Universal Robots URScript: T013_zai-org_GLM-4.7-FP8_edit_perf_rep1.urscript

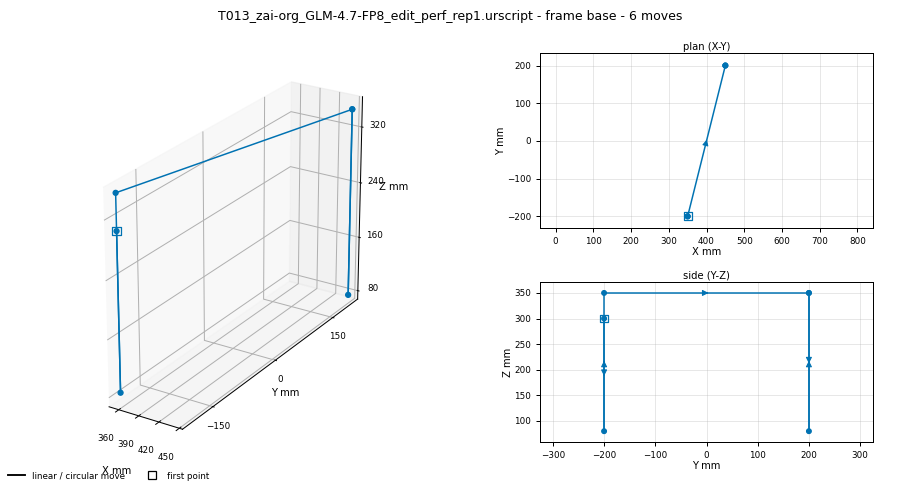
[picture p0: tool path of T013_zai-org_GLM-4.7-FP8_edit_perf_rep1.urscript in frame base, 6 of 8 moves have a stored position in this frame; points joined in program order, loops and branches not executed]
# Task: T013 — Collaborative suction palletizing — light boxes (Optimized)
# Generated by ENFIELD IR→URScript Translator
# Operating mode: collaborative | Max TCP speed: 0.250 m/s
# Robot: ur5e
#
# WARNING: This is auto-generated code for SIMULATION ONLY.
# Do NOT deploy to a physical robot without safety review.

def task_T013():
  # [0] E-Stop verify
  # E-Stop safety check (hardware-enforced on UR controller)
  if (get_digital_in(0) == True):
    popup("E-Stop active — aborting program.", error=True)
    halt
  end

  # [1] Home (Optimized: Increased joint velocity/acceleration)
  movej([0.0000, -1.5708, 1.5708, -1.5708, -1.5708, 0.0000], a=2.0000, v=1.5000)

  # [2] Above staging (Optimized: Max TCP speed, increased blend radius)
  movel(p[0.350000, -0.200000, 0.300000, 0.0000, 3.1416, 0.0000], a=1.2000, v=0.2500, r=0.0500)

  # [3] Descend to pick (Optimized: Slightly faster approach, no blend for precision)
  movel(p[0.350000, -0.200000, 0.080000, 0.0000, 3.1416, 0.0000], a=0.8000, v=0.1500, r=0.0000)

  # [4] Suction ON
  # set_tool (suction): {'vacuum_kpa': -40.0, 'state': 1.0}
  set_digital_out(0, True)

  # [5] Vacuum settle (Optimized: Reduced settle time for light payload)
  sleep(0.1000)

  # [6] Lift (Optimized: Max TCP speed, increased blend radius)
  movel(p[0.350000, -0.200000, 0.350000, 0.0000, 3.1416, 0.0000], a=1.2000, v=0.2500, r=0.0500)

  # [7] Transit to pallet (Optimized: Max TCP speed, increased blend radius)
  movel(p[0.450000, 0.200000, 0.350000, 0.0000, 3.1416, 0.0000], a=1.2000, v=0.2500, r=0.0500)

  # [8] Place on pallet (Optimized: Slightly faster approach, no blend for precision)
  movel(p[0.450000, 0.200000, 0.080000, 0.0000, 3.1416, 0.0000], a=0.8000, v=0.1500, r=0.0000)

  # [9] Suction OFF (Fixed: Corrected logic to False)
  # set_tool (suction): {'vacuum_kpa': 0.0, 'state': 0.0}
  set_digital_out(0, False)

  # [10] Release (Optimized: Reduced release time)
  sleep(0.1000)

  # [11] Retract (Optimized: Max TCP speed, increased blend radius)
  movel(p[0.450000, 0.200000, 0.350000, 0.0000, 3.1416, 0.0000], a=1.2000, v=0.2500, r=0.0500)

  # [12] Return home (Optimized: Increased joint velocity/acceleration)
  movej([0.0000, -1.5708, 1.5708, -1.5708, -1.5708, 0.0000], a=2.0000, v=1.5000)

end

# Entry point
task_T013()
